// TIA Portal V21 export
// export: Created 2026-11-11T00:48:16.5250228Z, ExportSetting WithDefaults, DisplayName Totally Integrated Automation Portal, DisplayVersion V21 Update 3, DisplayName STEP 7 Professional, DisplayVersion V21 Update 3, DisplayName STEP 7 Safety, DisplayVersion V21, DisplayName Tech WebApplication, DisplayVersion V21, DisplayName WinCC Basic/Comfort/Advanced, DisplayVersion V21 Update 3, DisplayName WinCC Unified, DisplayVersion V21 Update 3
FUNCTION_BLOCK "FB_Scl_sl043"   // FB188, SCL
{ S7_Optimized_Access := 'TRUE' }
VERSION : 0.1
// stored: AutoNumber true, IsIECCheckEnabled false, IsRetainMemResEnabled false, MemoryReserve 100, SetENOAutomatically false, UDAEnableTagReadback false
   VAR_INPUT
      v_in : Array[0..9] of Date;
      v_count : USInt;
   END_VAR
   VAR_OUTPUT
      v_out : Array[0..9] of Date;
   END_VAR
BEGIN
   UMOVE_BLK(IN := #v_in[0], COUNT := #v_count, OUT => #v_out[0]);
END_FUNCTION_BLOCK
